(* IEC 61131-3 sources: test/Class/HmiMemCircle, 1 file *)

(* ---- HmiMemCircle.st ---- *)
#include "..\..\Source\Common\hmi_nuc.h"

(*!
<Class
	Name               = "HmiMemCircle"
	Revision           = "0.0"
	RealtimeTask       = "false"
	CyclicTask         = "false"
	BackgroundTask     = "false"
	Sigmatek           = "true"
	OSInterface        = "false"
	HighPriority       = "false"
	Automatic          = "false"
	UpdateMode         = "Prescan"
	SharedCommandTable = "true"
	Objectsize         = "(284,120)">
	<Channels>
		<Server Name="ClassSvr" Visualized="false" Initialize="false" WriteProtected="true" Retentive="false"/>
		<Client Name="File" Required="true" Internal="false"/>
	</Channels>
	<Dependencies>
		<Files>
			<File Path=".\Source\Common\hmi_nuc.h" Include="true"/>
		</Files>
	</Dependencies>
</Class>
*)
HmiMemCircle : CLASS
  //Servers:
	ClassSvr 	: SvrChCmd_DINT;
  //Clients:
	File 	: CltChCmd_HmiFile;
  //Variables:
		Ptr 	: ^HMI_CTRL_CIRCLE;
		No 	: UDINT;
  //Functions:

	FUNCTION HmiMemCircle
		VAR_OUTPUT
			ret_code 	: ConfStates;
		END_VAR;

	FUNCTION GLOBAL Load
		VAR_OUTPUT
			retcode 	: BOOL;
		END_VAR;

	FUNCTION GLOBAL Free;

	FUNCTION HMI_CTRL_CIRCLE_Load
		VAR_INPUT
			tmp 	: ^HMI_CTRL_CIRCLE;
		END_VAR;

	FUNCTION GLOBAL Get
		VAR_INPUT
			index 	: UDINT;
		END_VAR
		VAR_OUTPUT
			retcode 	: ^HMI_CTRL_CIRCLE;
		END_VAR;
  //Tables:
	FUNCTION @STD
		VAR_OUTPUT
			ret_code	: CONFSTATES;
		END_VAR;
	FUNCTION GLOBAL TAB @CT_;
END_CLASS;

#pragma usingLtd HmiFile

FUNCTION HmiMemCircle::HmiMemCircle
	VAR_OUTPUT
		ret_code 	: ConfStates;
	END_VAR

  No  := 0;
  Ptr := NIL;
	ret_code := C_OK;

END_FUNCTION

FUNCTION HmiMemCircle::HMI_CTRL_CIRCLE_Load
	VAR_INPUT
		tmp 	: ^HMI_CTRL_CIRCLE;
	END_VAR

  File.Read_HMI_ROOM(#tmp^.room);
  File.FRead(#tmp^.color, 1);
  File.FRead(#tmp^.attrib, 4);
  File.Read_HMI_CHKBIT(#tmp^.chkbit);
  File.FRead(#tmp^.angle, 2);
  File.FRead(#tmp^.arc, 2);

END_FUNCTION

FUNCTION GLOBAL HmiMemCircle::Free
  var
    tmp : ^HMI_CTRL_CIRCLE;
  end_var

  tmp := Ptr;
  while(No) do
    No -= 1;
    free_HMI_CTRL_CIRCLE(tmp);
    tmp += sizeof(HMI_CTRL_CIRCLE);
  end_while;

  File.FMemory(#Ptr, 0);
  No  := 0;
  Ptr := NIL;

END_FUNCTION

FUNCTION GLOBAL HmiMemCircle::Load
	VAR_OUTPUT
		retcode 	: BOOL;
	END_VAR
  var
    anz : udint;
    ptmp : ^HMI_CTRL_CIRCLE;
  end_var;

  if(File.FRead(#anz, 4) = true) then
    if(File.FMemory(#Ptr$^void, anz * sizeof(HMI_CTRL_CIRCLE)) = true) then
      ptmp := Ptr;
      No   := anz;
      while(anz) do
        init_HMI_CTRL_CIRCLE(ptmp);
        HMI_CTRL_CIRCLE_Load(ptmp);
        ptmp += sizeof(HMI_CTRL_CIRCLE);
        anz  -= 1;
      end_while;
    end_if;
  end_if;

  retcode := File.FChkFile();
  ClassSvr := to_dint(No);

END_FUNCTION

FUNCTION GLOBAL HmiMemCircle::Get
	VAR_INPUT
		index 	: UDINT;
	END_VAR
	VAR_OUTPUT
		retcode 	: ^HMI_CTRL_CIRCLE;
	END_VAR

  retcode := NIL;
  if(index < No) then
    retcode := Ptr + (index * sizeof(HMI_CTRL_CIRCLE));
  end_if;

END_FUNCTION
